SUBAPPLICATION Uebung_155b (* Stoßfreie Hand/Auto-Umschaltung CTRL_PI_AR, realer Aufbau Pumpe + Durchflussmesser *)
  (* Standard: 61499-2; Description: Copyright (c) 2026 Meisterschulen am Ostbahnhof This program and the accompanying materials are made available under the terms of the Eclipse Public License 2.0 which is available at https://www.eclipse.org/legal/epl-2.0/ SPDX-License-Identifier: EPL-2.0 *)
  (* Version 1.0, 2026-11-15, Franz Höpfinger, Meisterschulen am Ostbahnhof, initial API and implementation and/or initial documentation *)
  PACKAGE Uebungen;
  IMPORT logiBUS::io::DI::logiBUS_DI::Input_I2;
  IMPORT logiBUS::io::DI::logiBUS_DI::Input_I3;
  IMPORT logiBUS::io::DI::logiBUS_DI::Input_I4;
  IMPORT logiBUS::io::DI::logiBUS_DI::Input_I5;
  IMPORT logiBUS::io::DI::logiBUS_DI::Input_I6;
  IMPORT logiBUS::io::DI::logiBUS_DI::Input_I7;
  IMPORT logiBUS::io::DI::logiBUS_DI::Input_I8;
  IMPORT logiBUS::io::DI::logiBUS_DI_Events::BUTTON_SINGLE_CLICK;
  IMPORT logiBUS::io::DQ::logiBUS_DO::Output_Q1;
  IMPORT logiBUS::io::PI::logiBUS_PI::PulseInput_I1;
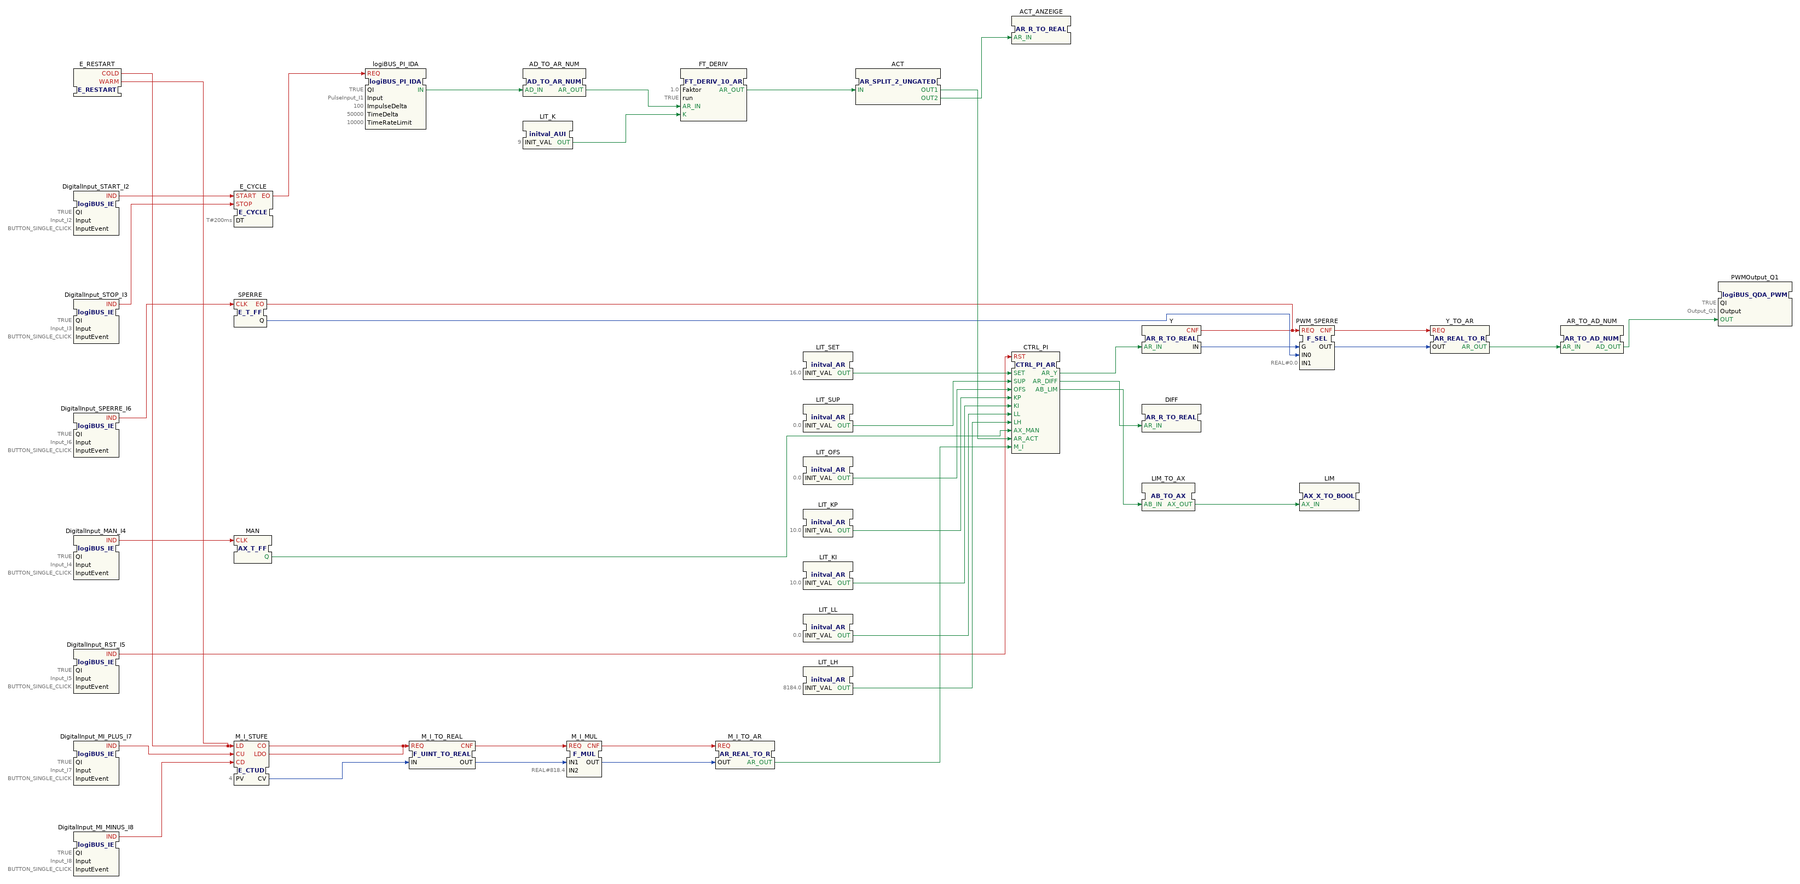
  (* Test stoßfreie Hand/Auto-Umschaltung (CTRL_PI_AR, OSCAT-Fix #385) Aufbau wie Übung 152: Durchflussmesser an I1, Pumpe an Q1. I2 = Takt starten, I3 = Takt stoppen. I4 = Hand/Auto (Start: Auto), I5 = RST Integrator, I6 = Pumpe sperren (PWM 0, Regler läuft weiter). Handwert M_I: Stufe 4 = 3273.6 (40 %); I7 +10 %, I8 -10 %. Watch: Y.IN, ACT_ANZEIGE.IN (Istwert), DIFF.IN, LIM.IN. 1) I4 Hand: Y = M_I. I4 Auto: Y springt nicht, regelt von M_I aus weiter. 2) Start in Auto: Y beginnt bei KP*DIFF (KP*DIFF), läuft nicht erst bis LH hoch. 3) Gegenprobe: in Auto I5 drücken -> Integrator 0, Y springt auf KP*DIFF. 4) Windup: I6 sperren -> Istwert fällt, Y läuft bis LH (8184), LIM = TRUE. Lösung im Projekt: RST bei steigender Freigabe. *)
  FBS
    CTRL_PI : OSCAT_adapter::Control::CTRL_PI_AR;
    LIT_SET : adapter::types::unidirectional::AR::initval::initval_AR(INIT_VAL := 16.0);
    LIT_SUP : adapter::types::unidirectional::AR::initval::initval_AR(INIT_VAL := 0.0);
    LIT_OFS : adapter::types::unidirectional::AR::initval::initval_AR(INIT_VAL := 0.0);
    LIT_KP : adapter::types::unidirectional::AR::initval::initval_AR(INIT_VAL := 10.0);
    LIT_KI : adapter::types::unidirectional::AR::initval::initval_AR(INIT_VAL := 10.0);
    LIT_LL : adapter::types::unidirectional::AR::initval::initval_AR(INIT_VAL := 0.0);
    LIT_LH : adapter::types::unidirectional::AR::initval::initval_AR(INIT_VAL := 8184.0);
    E_RESTART : iec61499::events::E_RESTART;
    SPERRE : iec61499::events::E_T_FF;
    MAN : adapter::events::unidirectional::AX_T_FF;
    Y : adapter::conversion::unidirectional::AR_R_TO_REAL;
    DIFF : adapter::conversion::unidirectional::AR_R_TO_REAL;
    LIM_TO_AX : adapter::conversion::unidirectional::AB_TO_AX;
    LIM : adapter::conversion::unidirectional::AX_X_TO_BOOL;
    DigitalInput_START_I2 : logiBUS::io::DI::logiBUS_IE(QI := TRUE, Input := Input_I2, InputEvent := BUTTON_SINGLE_CLICK);
    DigitalInput_STOP_I3 : logiBUS::io::DI::logiBUS_IE(QI := TRUE, Input := Input_I3, InputEvent := BUTTON_SINGLE_CLICK);
    E_CYCLE : iec61499::events::E_CYCLE(DT := T#200ms);
    logiBUS_PI_IDA : logiBUS::io::PI::logiBUS_PI_IDA(QI := TRUE, Input := PulseInput_I1, ImpulseDelta := 100, TimeDelta := 50000, TimeRateLimit := 10000);
    AD_TO_AR_NUM : adapter::conversion::unidirectional::AD_TO_AR_NUM;
    FT_DERIV : OSCAT_adapter::Control::FT_DERIV_10_AR(Faktor := 1.0, run := TRUE);
    LIT_K : adapter::types::unidirectional::AUI::initval::initval_AUI(INIT_VAL := 9);
    ACT : adapter::events::unidirectional::AR_SPLIT_2_UNGATED;
    ACT_ANZEIGE : adapter::conversion::unidirectional::AR_R_TO_REAL;
    DigitalInput_MAN_I4 : logiBUS::io::DI::logiBUS_IE(QI := TRUE, Input := Input_I4, InputEvent := BUTTON_SINGLE_CLICK);
    DigitalInput_RST_I5 : logiBUS::io::DI::logiBUS_IE(QI := TRUE, Input := Input_I5, InputEvent := BUTTON_SINGLE_CLICK);
    DigitalInput_SPERRE_I6 : logiBUS::io::DI::logiBUS_IE(QI := TRUE, Input := Input_I6, InputEvent := BUTTON_SINGLE_CLICK);
    DigitalInput_MI_PLUS_I7 : logiBUS::io::DI::logiBUS_IE(QI := TRUE, Input := Input_I7, InputEvent := BUTTON_SINGLE_CLICK);
    DigitalInput_MI_MINUS_I8 : logiBUS::io::DI::logiBUS_IE(QI := TRUE, Input := Input_I8, InputEvent := BUTTON_SINGLE_CLICK);
    M_I_STUFE : iec61499::events::E_CTUD(PV := 4);
    M_I_TO_REAL : iec61131::conversion::F_UINT_TO_REAL;
    M_I_MUL : iec61131::arithmetic::F_MUL(IN2 := REAL#818.4);
    M_I_TO_AR : adapter::conversion::unidirectional::AR_REAL_TO_R;
    PWM_SPERRE : iec61131::selection::F_SEL(IN1 := REAL#0.0);
    Y_TO_AR : adapter::conversion::unidirectional::AR_REAL_TO_R;
    AR_TO_AD_NUM : adapter::conversion::unidirectional::AR_TO_AD_NUM;
    PWMOutput_Q1 : logiBUS::io::DQ::logiBUS_QDA_PWM(QI := TRUE, Output := Output_Q1);
  END_FBS
  EVENT_CONNECTIONS
    DigitalInput_START_I2.IND TO E_CYCLE.START;
    DigitalInput_STOP_I3.IND TO E_CYCLE.STOP;
    E_CYCLE.EO TO logiBUS_PI_IDA.REQ;
    DigitalInput_MAN_I4.IND TO MAN.CLK;
    DigitalInput_RST_I5.IND TO CTRL_PI.RST;
    DigitalInput_SPERRE_I6.IND TO SPERRE.CLK;
    E_RESTART.COLD TO M_I_STUFE.LD;
    E_RESTART.WARM TO M_I_STUFE.LD;
    DigitalInput_MI_PLUS_I7.IND TO M_I_STUFE.CU;
    DigitalInput_MI_MINUS_I8.IND TO M_I_STUFE.CD;
    M_I_STUFE.CO TO M_I_TO_REAL.REQ;
    M_I_STUFE.LDO TO M_I_TO_REAL.REQ;
    M_I_TO_REAL.CNF TO M_I_MUL.REQ;
    M_I_MUL.CNF TO M_I_TO_AR.REQ;
    Y.CNF TO PWM_SPERRE.REQ;
    SPERRE.EO TO PWM_SPERRE.REQ;
    PWM_SPERRE.CNF TO Y_TO_AR.REQ;
  END_CONNECTIONS
  DATA_CONNECTIONS
    M_I_STUFE.CV TO M_I_TO_REAL.IN;
    M_I_TO_REAL.OUT TO M_I_MUL.IN1;
    M_I_MUL.OUT TO M_I_TO_AR.OUT;
    SPERRE.Q TO PWM_SPERRE.G;
    Y.IN TO PWM_SPERRE.IN0;
    PWM_SPERRE.OUT TO Y_TO_AR.OUT;
  END_CONNECTIONS
  ADAPTER_CONNECTIONS
    LIT_SET.OUT TO CTRL_PI.SET;
    LIT_SUP.OUT TO CTRL_PI.SUP;
    LIT_OFS.OUT TO CTRL_PI.OFS;
    LIT_KP.OUT TO CTRL_PI.KP;
    LIT_KI.OUT TO CTRL_PI.KI;
    LIT_LL.OUT TO CTRL_PI.LL;
    LIT_LH.OUT TO CTRL_PI.LH;
    MAN.Q TO CTRL_PI.AX_MAN;
    CTRL_PI.AR_Y TO Y.AR_IN;
    CTRL_PI.AR_DIFF TO DIFF.AR_IN;
    CTRL_PI.AB_LIM TO LIM_TO_AX.AB_IN;
    LIM_TO_AX.AX_OUT TO LIM.AX_IN;
    logiBUS_PI_IDA.IN TO AD_TO_AR_NUM.AD_IN;
    AD_TO_AR_NUM.AR_OUT TO FT_DERIV.AR_IN;
    LIT_K.OUT TO FT_DERIV.K;
    FT_DERIV.AR_OUT TO ACT.IN;
    ACT.OUT1 TO CTRL_PI.AR_ACT;
    ACT.OUT2 TO ACT_ANZEIGE.AR_IN;
    M_I_TO_AR.AR_OUT TO CTRL_PI.M_I;
    Y_TO_AR.AR_OUT TO AR_TO_AD_NUM.AR_IN;
    AR_TO_AD_NUM.AD_OUT TO PWMOutput_Q1.OUT;
  END_CONNECTIONS
END_SUBAPPLICATION
